(* IEC 61131-3 sources: BODAS-RC27-18_40/st/bodas_rc18_12_27_18_40/plc_logic/application/dsm_easyconfig/structure (part 3) *)

(* ---- dfc_rbr_outa09ot-DFC_rbr_outA09OT.st ---- *)
(* --- Interface --- *)
{attribute 'external_name' := 'cmp_rts_DFC_rbr_outA09OT'}
TYPE DFC_rbr_outA09OT :
STRUCT
	DTC: UDINT := 16#142D00;
	DFCid: UINT := 305;
	debounceMethod: USINT := TIME_UP_DOWN;
END_STRUCT
END_TYPE

(* ---- dfc_rbr_outa09scb-DFC_rbr_outA09SCB.st ---- *)
(* --- Interface --- *)
{attribute 'external_name' := 'cmp_rts_DFC_rbr_outA09SCB'}
TYPE DFC_rbr_outA09SCB :
STRUCT
	DTC: UDINT := 16#142E00;
	DFCid: UINT := 306;
	debounceMethod: USINT := TIME_UP_DOWN;
END_STRUCT
END_TYPE

(* ---- dfc_rbr_outa09scg-DFC_rbr_outA09SCG.st ---- *)
(* --- Interface --- *)
{attribute 'external_name' := 'cmp_rts_DFC_rbr_outA09SCG'}
TYPE DFC_rbr_outA09SCG :
STRUCT
	DTC: UDINT := 16#142F00;
	DFCid: UINT := 307;
	debounceMethod: USINT := TIME_UP_DOWN;
END_STRUCT
END_TYPE

(* ---- dfc_rbr_outa09unintended-DFC_rbr_outA09Unintended.st ---- *)
(* --- Interface --- *)
{attribute 'external_name' := 'cmp_rts_DFC_rbr_outA09Unintended'}
TYPE DFC_rbr_outA09Unintended :
STRUCT
	DTC: UDINT := 16#14B900;
	DFCid: UINT := 680;
	debounceMethod: USINT := NO_DEBOUNCE;
END_STRUCT
END_TYPE

(* ---- dfc_rbr_outa10oc-DFC_rbr_outA10OC.st ---- *)
(* --- Interface --- *)
{attribute 'external_name' := 'cmp_rts_DFC_rbr_outA10OC'}
TYPE DFC_rbr_outA10OC :
STRUCT
	DTC: UDINT := 16#143000;
	DFCid: UINT := 681;
	debounceMethod: USINT := NO_DEBOUNCE;
END_STRUCT
END_TYPE

(* ---- dfc_rbr_outa10ol-DFC_rbr_outA10OL.st ---- *)
(* --- Interface --- *)
{attribute 'external_name' := 'cmp_rts_DFC_rbr_outA10OL'}
TYPE DFC_rbr_outA10OL :
STRUCT
	DTC: UDINT := 16#143100;
	DFCid: UINT := 308;
	debounceMethod: USINT := TIME_UP_DOWN;
END_STRUCT
END_TYPE

(* ---- dfc_rbr_outa10ot-DFC_rbr_outA10OT.st ---- *)
(* --- Interface --- *)
{attribute 'external_name' := 'cmp_rts_DFC_rbr_outA10OT'}
TYPE DFC_rbr_outA10OT :
STRUCT
	DTC: UDINT := 16#143200;
	DFCid: UINT := 309;
	debounceMethod: USINT := TIME_UP_DOWN;
END_STRUCT
END_TYPE

(* ---- dfc_rbr_outa10scb-DFC_rbr_outA10SCB.st ---- *)
(* --- Interface --- *)
{attribute 'external_name' := 'cmp_rts_DFC_rbr_outA10SCB'}
TYPE DFC_rbr_outA10SCB :
STRUCT
	DTC: UDINT := 16#143300;
	DFCid: UINT := 310;
	debounceMethod: USINT := TIME_UP_DOWN;
END_STRUCT
END_TYPE

(* ---- dfc_rbr_outa10scg-DFC_rbr_outA10SCG.st ---- *)
(* --- Interface --- *)
{attribute 'external_name' := 'cmp_rts_DFC_rbr_outA10SCG'}
TYPE DFC_rbr_outA10SCG :
STRUCT
	DTC: UDINT := 16#143400;
	DFCid: UINT := 311;
	debounceMethod: USINT := TIME_UP_DOWN;
END_STRUCT
END_TYPE

(* ---- dfc_rbr_outa10unintended-DFC_rbr_outA10Unintended.st ---- *)
(* --- Interface --- *)
{attribute 'external_name' := 'cmp_rts_DFC_rbr_outA10Unintended'}
TYPE DFC_rbr_outA10Unintended :
STRUCT
	DTC: UDINT := 16#14BA00;
	DFCid: UINT := 682;
	debounceMethod: USINT := NO_DEBOUNCE;
END_STRUCT
END_TYPE

(* ---- dfc_rbr_outa11ol-DFC_rbr_outA11OL.st ---- *)
(* --- Interface --- *)
{attribute 'external_name' := 'cmp_rts_DFC_rbr_outA11OL'}
TYPE DFC_rbr_outA11OL :
STRUCT
	DTC: UDINT := 16#143500;
	DFCid: UINT := 312;
	debounceMethod: USINT := TIME_UP_DOWN;
END_STRUCT
END_TYPE

(* ---- dfc_rbr_outa11ot-DFC_rbr_outA11OT.st ---- *)
(* --- Interface --- *)
{attribute 'external_name' := 'cmp_rts_DFC_rbr_outA11OT'}
TYPE DFC_rbr_outA11OT :
STRUCT
	DTC: UDINT := 16#143600;
	DFCid: UINT := 313;
	debounceMethod: USINT := TIME_UP_DOWN;
END_STRUCT
END_TYPE

(* ---- dfc_rbr_outa11scb-DFC_rbr_outA11SCB.st ---- *)
(* --- Interface --- *)
{attribute 'external_name' := 'cmp_rts_DFC_rbr_outA11SCB'}
TYPE DFC_rbr_outA11SCB :
STRUCT
	DTC: UDINT := 16#143700;
	DFCid: UINT := 314;
	debounceMethod: USINT := TIME_UP_DOWN;
END_STRUCT
END_TYPE

(* ---- dfc_rbr_outa11scg-DFC_rbr_outA11SCG.st ---- *)
(* --- Interface --- *)
{attribute 'external_name' := 'cmp_rts_DFC_rbr_outA11SCG'}
TYPE DFC_rbr_outA11SCG :
STRUCT
	DTC: UDINT := 16#143800;
	DFCid: UINT := 315;
	debounceMethod: USINT := TIME_UP_DOWN;
END_STRUCT
END_TYPE

(* ---- dfc_rbr_outa12or-DFC_rbr_outA12OR.st ---- *)
(* --- Interface --- *)
{attribute 'external_name' := 'cmp_rts_DFC_rbr_outA12OR'}
TYPE DFC_rbr_outA12OR :
STRUCT
	DTC: UDINT := 16#143900;
	DFCid: UINT := 316;
	debounceMethod: USINT := TIME_UP_DOWN;
END_STRUCT
END_TYPE

(* ---- dfc_rbr_outa12scb-DFC_rbr_outA12SCB.st ---- *)
(* --- Interface --- *)
{attribute 'external_name' := 'cmp_rts_DFC_rbr_outA12SCB'}
TYPE DFC_rbr_outA12SCB :
STRUCT
	DTC: UDINT := 16#143A00;
	DFCid: UINT := 317;
	debounceMethod: USINT := TIME_UP_DOWN;
END_STRUCT
END_TYPE

(* ---- dfc_rbr_outa12scg-DFC_rbr_outA12SCG.st ---- *)
(* --- Interface --- *)
{attribute 'external_name' := 'cmp_rts_DFC_rbr_outA12SCG'}
TYPE DFC_rbr_outA12SCG :
STRUCT
	DTC: UDINT := 16#143B00;
	DFCid: UINT := 318;
	debounceMethod: USINT := TIME_UP_DOWN;
END_STRUCT
END_TYPE

(* ---- dfc_rbr_outa16ol-DFC_rbr_outA16OL.st ---- *)
(* --- Interface --- *)
{attribute 'external_name' := 'cmp_rts_DFC_rbr_outA16OL'}
TYPE DFC_rbr_outA16OL :
STRUCT
	DTC: UDINT := 16#143C00;
	DFCid: UINT := 319;
	debounceMethod: USINT := TIME_UP_DOWN;
END_STRUCT
END_TYPE

(* ---- dfc_rbr_outa16ot-DFC_rbr_outA16OT.st ---- *)
(* --- Interface --- *)
{attribute 'external_name' := 'cmp_rts_DFC_rbr_outA16OT'}
TYPE DFC_rbr_outA16OT :
STRUCT
	DTC: UDINT := 16#143D00;
	DFCid: UINT := 320;
	debounceMethod: USINT := TIME_UP_DOWN;
END_STRUCT
END_TYPE

(* ---- dfc_rbr_outa16scb-DFC_rbr_outA16SCB.st ---- *)
(* --- Interface --- *)
{attribute 'external_name' := 'cmp_rts_DFC_rbr_outA16SCB'}
TYPE DFC_rbr_outA16SCB :
STRUCT
	DTC: UDINT := 16#143E00;
	DFCid: UINT := 321;
	debounceMethod: USINT := TIME_UP_DOWN;
END_STRUCT
END_TYPE

(* ---- dfc_rbr_outa16scg-DFC_rbr_outA16SCG.st ---- *)
(* --- Interface --- *)
{attribute 'external_name' := 'cmp_rts_DFC_rbr_outA16SCG'}
TYPE DFC_rbr_outA16SCG :
STRUCT
	DTC: UDINT := 16#143F00;
	DFCid: UINT := 322;
	debounceMethod: USINT := TIME_UP_DOWN;
END_STRUCT
END_TYPE

(* ---- dfc_rbr_outa17oc-DFC_rbr_outA17OC.st ---- *)
(* --- Interface --- *)
{attribute 'external_name' := 'cmp_rts_DFC_rbr_outA17OC'}
TYPE DFC_rbr_outA17OC :
STRUCT
	DTC: UDINT := 16#144000;
	DFCid: UINT := 683;
	debounceMethod: USINT := NO_DEBOUNCE;
END_STRUCT
END_TYPE

(* ---- dfc_rbr_outa17ol-DFC_rbr_outA17OL.st ---- *)
(* --- Interface --- *)
{attribute 'external_name' := 'cmp_rts_DFC_rbr_outA17OL'}
TYPE DFC_rbr_outA17OL :
STRUCT
	DTC: UDINT := 16#144100;
	DFCid: UINT := 323;
	debounceMethod: USINT := TIME_UP_DOWN;
END_STRUCT
END_TYPE

(* ---- dfc_rbr_outa17or-DFC_rbr_outA17OR.st ---- *)
(* --- Interface --- *)
{attribute 'external_name' := 'cmp_rts_DFC_rbr_outA17OR'}
TYPE DFC_rbr_outA17OR :
STRUCT
	DTC: UDINT := 16#144200;
	DFCid: UINT := 324;
	debounceMethod: USINT := TIME_UP_DOWN;
END_STRUCT
END_TYPE

(* ---- dfc_rbr_outa17ot-DFC_rbr_outA17OT.st ---- *)
(* --- Interface --- *)
{attribute 'external_name' := 'cmp_rts_DFC_rbr_outA17OT'}
TYPE DFC_rbr_outA17OT :
STRUCT
	DTC: UDINT := 16#144300;
	DFCid: UINT := 325;
	debounceMethod: USINT := TIME_UP_DOWN;
END_STRUCT
END_TYPE

(* ---- dfc_rbr_outa17scb-DFC_rbr_outA17SCB.st ---- *)
(* --- Interface --- *)
{attribute 'external_name' := 'cmp_rts_DFC_rbr_outA17SCB'}
TYPE DFC_rbr_outA17SCB :
STRUCT
	DTC: UDINT := 16#144400;
	DFCid: UINT := 326;
	debounceMethod: USINT := TIME_UP_DOWN;
END_STRUCT
END_TYPE

(* ---- dfc_rbr_outa17scg-DFC_rbr_outA17SCG.st ---- *)
(* --- Interface --- *)
{attribute 'external_name' := 'cmp_rts_DFC_rbr_outA17SCG'}
TYPE DFC_rbr_outA17SCG :
STRUCT
	DTC: UDINT := 16#144500;
	DFCid: UINT := 327;
	debounceMethod: USINT := TIME_UP_DOWN;
END_STRUCT
END_TYPE

(* ---- dfc_rbr_outa17unintended-DFC_rbr_outA17Unintended.st ---- *)
(* --- Interface --- *)
{attribute 'external_name' := 'cmp_rts_DFC_rbr_outA17Unintended'}
TYPE DFC_rbr_outA17Unintended :
STRUCT
	DTC: UDINT := 16#14BB00;
	DFCid: UINT := 684;
	debounceMethod: USINT := NO_DEBOUNCE;
END_STRUCT
END_TYPE

(* ---- dfc_rbr_outa18oc-DFC_rbr_outA18OC.st ---- *)
(* --- Interface --- *)
{attribute 'external_name' := 'cmp_rts_DFC_rbr_outA18OC'}
TYPE DFC_rbr_outA18OC :
STRUCT
	DTC: UDINT := 16#144600;
	DFCid: UINT := 685;
	debounceMethod: USINT := NO_DEBOUNCE;
END_STRUCT
END_TYPE

(* ---- dfc_rbr_outa18ol-DFC_rbr_outA18OL.st ---- *)
(* --- Interface --- *)
{attribute 'external_name' := 'cmp_rts_DFC_rbr_outA18OL'}
TYPE DFC_rbr_outA18OL :
STRUCT
	DTC: UDINT := 16#144700;
	DFCid: UINT := 328;
	debounceMethod: USINT := TIME_UP_DOWN;
END_STRUCT
END_TYPE

(* ---- dfc_rbr_outa18ot-DFC_rbr_outA18OT.st ---- *)
(* --- Interface --- *)
{attribute 'external_name' := 'cmp_rts_DFC_rbr_outA18OT'}
TYPE DFC_rbr_outA18OT :
STRUCT
	DTC: UDINT := 16#144800;
	DFCid: UINT := 329;
	debounceMethod: USINT := TIME_UP_DOWN;
END_STRUCT
END_TYPE

(* ---- dfc_rbr_outa18scb-DFC_rbr_outA18SCB.st ---- *)
(* --- Interface --- *)
{attribute 'external_name' := 'cmp_rts_DFC_rbr_outA18SCB'}
TYPE DFC_rbr_outA18SCB :
STRUCT
	DTC: UDINT := 16#144900;
	DFCid: UINT := 330;
	debounceMethod: USINT := TIME_UP_DOWN;
END_STRUCT
END_TYPE

(* ---- dfc_rbr_outa18scg-DFC_rbr_outA18SCG.st ---- *)
(* --- Interface --- *)
{attribute 'external_name' := 'cmp_rts_DFC_rbr_outA18SCG'}
TYPE DFC_rbr_outA18SCG :
STRUCT
	DTC: UDINT := 16#144A00;
	DFCid: UINT := 331;
	debounceMethod: USINT := TIME_UP_DOWN;
END_STRUCT
END_TYPE

(* ---- dfc_rbr_outa18unintended-DFC_rbr_outA18Unintended.st ---- *)
(* --- Interface --- *)
{attribute 'external_name' := 'cmp_rts_DFC_rbr_outA18Unintended'}
TYPE DFC_rbr_outA18Unintended :
STRUCT
	DTC: UDINT := 16#14BC00;
	DFCid: UINT := 686;
	debounceMethod: USINT := NO_DEBOUNCE;
END_STRUCT
END_TYPE

(* ---- dfc_rbr_outa19oc-DFC_rbr_outA19OC.st ---- *)
(* --- Interface --- *)
{attribute 'external_name' := 'cmp_rts_DFC_rbr_outA19OC'}
TYPE DFC_rbr_outA19OC :
STRUCT
	DTC: UDINT := 16#144B00;
	DFCid: UINT := 687;
	debounceMethod: USINT := NO_DEBOUNCE;
END_STRUCT
END_TYPE

(* ---- dfc_rbr_outa19ol-DFC_rbr_outA19OL.st ---- *)
(* --- Interface --- *)
{attribute 'external_name' := 'cmp_rts_DFC_rbr_outA19OL'}
TYPE DFC_rbr_outA19OL :
STRUCT
	DTC: UDINT := 16#144C00;
	DFCid: UINT := 332;
	debounceMethod: USINT := TIME_UP_DOWN;
END_STRUCT
END_TYPE

(* ---- dfc_rbr_outa19or-DFC_rbr_outA19OR.st ---- *)
(* --- Interface --- *)
{attribute 'external_name' := 'cmp_rts_DFC_rbr_outA19OR'}
TYPE DFC_rbr_outA19OR :
STRUCT
	DTC: UDINT := 16#144D00;
	DFCid: UINT := 333;
	debounceMethod: USINT := TIME_UP_DOWN;
END_STRUCT
END_TYPE
